(* IEC 61131-3 sources: axsharp/src/AXSharp.compiler/tests/AXSharp.CompilerTests/samples/plt/lib/test, 1 file *)

(* ---- test.st ---- *)
USING AxUnit;
USING MyLibrary;

NAMESPACE MyTest

    {TestFixture}
    CLASS MyTestFixture

        VAR PROTECTED
            testInstance : MyClass;
        END_VAR

        {Test}
        METHOD PUBLIC MyTestMethod
            VAR_TEMP
                result : BOOL;
            END_VAR

            result := testInstance.MyMethod();

            Assert.Equal(actual := result, expected := FALSE);

        END_METHOD
    END_CLASS

END_NAMESPACE
